(* IEC 61131-3 sources: s7-to-codesys/src/POUs/S7Compat/F_S5Update, 2 files *)

(* ---- F_S5Update.decl.st ---- *)
// Назначение: пересчёт таймера S5 на текущий момент F_S7Now(): у идущего таймера — остаток, по истечении
//             времени — останов и состояние Q по виду пуска (SD, SS — TRUE; SP, SE, SF — FALSE). Возвращает
//             остаток. Его вызывают все функции, которые читают таймер или останавливают его: в S7 время
//             уменьшает часовой процесс CPU асинхронно циклу, и опрос видит состояние на момент чтения.
//             Разность моментов — по модулю 2^32 (переход TIME через ноль переносится).
// Автор:      kr0nsch
// Версия:     1.2.0
// Документ:   docs/MAPPING_STL.md, правило s5.timebase; docs/ASSUMPTIONS.md, запись L13
FUNCTION F_S5Update : TIME
VAR_IN_OUT
    stTimer : ST_S5Timer;   // таймер
END_VAR
VAR
    tElapsed : TIME;        // прошло с пуска
END_VAR

(* ---- F_S5Update.impl.st ---- *)
IF stTimer.xRunning THEN
    tElapsed := F_S7Now() - stTimer.tStart;
    IF tElapsed >= stTimer.tPreset THEN
        stTimer.xRunning := FALSE;
        stTimer.xQ := stTimer.xQAtEnd;
        stTimer.tRest := T#0MS;
    ELSE
        stTimer.tRest := stTimer.tPreset - tElapsed;
    END_IF
END_IF
F_S5Update := stTimer.tRest;
